// TIA Portal V17 export
// export: Created 2026-09-23T08:10:24.1555226Z, ExportSetting None, DisplayName Totally Integrated Automation Portal, DisplayVersion V17, DisplayName TIA Portal Openness, DisplayVersion V17, DisplayName TIA Portal Version Control Interface, DisplayVersion V17, DisplayName STEP 7 Professional, DisplayVersion V17, DisplayName STEP 7 Safety, DisplayVersion V17, DisplayName WinCC Advanced, DisplayVersion V17
DATA_BLOCK "AnimationTimer"   // DB1
{ S7_Optimized_Access := 'FALSE' }
   VAR
      T1 : TON_TIME;
      T2 : TON_TIME;
      T3 : TON_TIME;
      T4 : TON_TIME;
   END_VAR
BEGIN
END_DATA_BLOCK
